(* CODESYS project qualified_candidate.project

Project tree, tasks and I/O mapping:
  PLCWinNT : CODESYS Control Win V3 x64, CODESYS, version 3.5.22.40
    application Application
      libraries: Standard, * (System)
      task MainTask (cyclic, interval t#50ms, priority 1) calls PLC_PRG
      program PLC_PRG [ST]
*)

// PLCWinNT/Application/PLC_PRG
PROGRAM PLC_PRG
VAR
END_VAR

;

END_PROGRAM
